(* IEC 61131-3 sources: Jacob-Formschaumtechnik-ISEL-CNC-Retrofit/twincat/PLC/src/4_Machine, 9 files *)

(* ---- FB_Homing.st ---- *)
(* Referenzfahrt als Ablauf: Z zuerst (Spindel nach oben), dann Querachse, dann Portal (Gantry).
   Reihenfolge und Richtung einstellbar (Anforderung 2.2.1). Der Baustein fordert die Fahrt an,
   die Bewegung selbst macht die CNC bzw. der Antrieb. Gantry-Ausrichtung beider Portalseiten
   gehoert in die CNC-Parametrierung. Gruppen: 1 = Z, 2 = X (Quer), 3 = Y (Portal).
   [Annahme] Reihenfolge Z, X, Y, bis Maschinenaufbau bestaetigt.
   Befund 8: Je Gruppe ein Handshake. Erst kommt ein Ruecksetz-Impuls (aResetHomed), dann muss aHomed
   FALSE werden, danach steht bHomeCmd als Pegel, bis aHomed wieder TRUE ist. Zwischen zwei Gruppen
   faellt bHomeCmd mindestens einen Zyklus. Einzelne X/Y-Referenzfahrt nur mit referenziertem Z. *)
FUNCTION_BLOCK FB_Homing
VAR_INPUT
    bStart       : BOOL;                      (* Impuls: alle Achsen in Reihenfolge *)
    aStartAxis   : ARRAY[1..3] OF BOOL;       (* Impuls: nur diese Gruppe *)
    bAbort       : BOOL;
    bHomingOk    : BOOL;
    aHomed       : ARRAY[1..3] OF BOOL;       (* je Gruppe, aus dem einheitlichen Referenzstatus *)
    aOrder       : ARRAY[1..3] OF USINT := [1, 2, 3];
    tTimeout     : TIME := T#120S;
END_VAR
VAR_OUTPUT
    bBusy        : BOOL;
    bDone        : BOOL;
    bError       : BOOL;
    nActiveGroup : USINT;                     (* Gruppe, die gerade referenziert wird, 0 = keine *)
    bHomeCmd     : BOOL;                      (* Anforderung an die CNC/den Antrieb fuer nActiveGroup *)
    aResetHomed  : ARRAY[1..3] OF BOOL;       (* Impuls: Referenzstatus dieser Gruppe loeschen *)
    eHomeState   : ARRAY[1..3] OF E_HomeState;
    nStepOut     : USINT;
END_VAR
VAR
    nStep      : INT;
    nSub       : INT;                         (* 0 Reset senden, 1 auf Reset warten, 2 fahren *)
    nSingle    : USINT;
    rtStart    : R_TRIG;
    rtSingle   : ARRAY[1..3] OF R_TRIG;
    tonTimeout : TON;
    i          : INT;
END_VAR

rtStart(CLK := bStart);
FOR i := 1 TO 3 DO
    rtSingle[i](CLK := aStartAxis[i]);
    aResetHomed[i] := FALSE;
END_FOR
bHomeCmd := FALSE;

IF bAbort OR (bBusy AND NOT bHomingOk) THEN
    IF bBusy AND nActiveGroup > 0 THEN eHomeState[nActiveGroup] := E_HomeState.Open; END_IF
    nStep := 0; nSub := 0; bBusy := FALSE; nActiveGroup := 0; tonTimeout(IN := FALSE);
END_IF

CASE nStep OF
    0:
        IF bHomingOk THEN
            IF rtStart.Q THEN
                bDone := FALSE; bError := FALSE; bBusy := TRUE; nSingle := 0; nStep := 1; nSub := 0;
                FOR i := 1 TO 3 DO eHomeState[i] := E_HomeState.Open; END_FOR
            ELSE
                FOR i := 1 TO 3 DO
                    IF rtSingle[i].Q AND NOT bBusy THEN
                        IF i > 1 AND NOT aHomed[1] THEN
                            bError := TRUE;    (* Z muss zuerst referenziert sein *)
                        ELSE
                            bDone := FALSE; bError := FALSE; bBusy := TRUE; nSingle := TO_USINT(i);
                            nStep := 1; nSub := 0;
                            eHomeState[i] := E_HomeState.Open;
                        END_IF
                    END_IF
                END_FOR
            END_IF
        END_IF
    1, 2, 3:
        IF nSingle > 0 THEN
            nActiveGroup := nSingle;
        ELSE
            nActiveGroup := aOrder[nStep];
        END_IF
        tonTimeout(IN := TRUE, PT := tTimeout);
        CASE nSub OF
            0:  aResetHomed[nActiveGroup] := TRUE;
                eHomeState[nActiveGroup] := E_HomeState.Running;
                nSub := 1;
            1:  IF NOT aHomed[nActiveGroup] THEN nSub := 2; END_IF
            2:  bHomeCmd := TRUE;
                IF aHomed[nActiveGroup] THEN
                    eHomeState[nActiveGroup] := E_HomeState.Done;
                    tonTimeout(IN := FALSE);
                    nSub := 0;
                    IF nSingle > 0 THEN nStep := 4; ELSE nStep := nStep + 1; END_IF
                END_IF
        END_CASE
        IF tonTimeout.Q THEN
            eHomeState[nActiveGroup] := E_HomeState.Error;
            bError := TRUE; bBusy := FALSE; nActiveGroup := 0; nStep := 0; nSub := 0;
            tonTimeout(IN := FALSE);
        END_IF
    4:
        bDone := TRUE; bBusy := FALSE; nActiveGroup := 0; nStep := 0; nSub := 0;
END_CASE
nStepOut := TO_USINT(nStep);
END_FUNCTION_BLOCK

(* ---- FB_Interlocks.st ---- *)
(* Verriegelungsmatrix. Reine Logik ohne Hardwarebezug, daher voll testbar.
   Jede Zeile haengt an einer Anforderung aus der Funktionsliste (Platzhalter-IDs bis Lastenheft da ist). *)
FUNCTION_BLOCK FB_Interlocks
VAR_INPUT
    eMode          : E_OpMode;
    eState         : E_MachState;
    bSafetyOk      : BOOL;
    bAllHomed      : BOOL;
    bDrivesEnabled : BOOL;
    bHmiLinkOk     : BOOL;
    bAnyR2OrHigher : BOOL;
    bAnyR3OrHigher : BOOL;
    bAirOk         : BOOL;
    bHomingBusy    : BOOL;      (* Referenzfahrt laeuft (Befund 8c) *)
    bLimitFreeRun  : BOOL;      (* nur Endschalter-R3 aktiv, Freifahren erlaubt (Befund 15) *)
END_VAR
VAR_OUTPUT
    bProgramStartOk : BOOL;   (* Auto: Start erlaubt *)
    bJogOk          : BOOL;   (* Tippen erlaubt *)
    bHomingOk       : BOOL;
    bSpindleOk      : BOOL;   (* Spindel darf laufen *)
    bAuxOk          : BOOL;   (* Absaugung, Blasluft, Vakuum von Hand *)
    bModeChangeOk   : BOOL;   (* Wechsel nur ohne aktives Programm *)
END_VAR

bProgramStartOk := eMode = E_OpMode.Auto OR eMode = E_OpMode.Setup;
bProgramStartOk := bProgramStartOk AND bSafetyOk AND bDrivesEnabled AND bAllHomed
                   AND NOT bAnyR2OrHigher AND bAirOk AND eState <> E_MachState.Execute AND NOT bHomingBusy;

bJogOk := eMode = E_OpMode.Hand AND bSafetyOk AND bDrivesEnabled AND bHmiLinkOk
          AND (NOT bAnyR3OrHigher OR bLimitFreeRun) AND eState <> E_MachState.Execute AND NOT bHomingBusy;

(* Referenzfahrt nur in Hand und nur im Zustand Idle (nicht in Held/Execute) *)
bHomingOk := eMode = E_OpMode.Hand AND bSafetyOk AND bDrivesEnabled AND NOT bAnyR3OrHigher AND eState = E_MachState.Idle;

bSpindleOk := bSafetyOk AND NOT bAnyR3OrHigher AND eMode <> E_OpMode.Setup;

bAuxOk := bSafetyOk AND eState <> E_MachState.EStop;

bModeChangeOk := eState <> E_MachState.Execute AND eState <> E_MachState.Held;
END_FUNCTION_BLOCK

(* ---- FB_Jog.st ---- *)
(* Tippbetrieb aus der HMI (Anforderungen 2.3.1 und 2.3.2). Nur mit Lebenszeichen der HMI, nur
   in Betriebsart Hand. Befund 6 der Papierpruefung: Tippen startet nur mit einer steigenden Flanke
   der Taste, waehrend alle Freigaben bestehen. Eine beim Wiederkehren der Freigabe (Quittierung,
   Sicherheitskreis, HMI-Lebenszeichen) noch gehaltene Taste startet nichts. Die Achsnummer wird
   beim Start festgehalten. Die Bewegung selbst fordert die CNC an. *)
FUNCTION_BLOCK FB_Jog
VAR_INPUT
    bJogOk       : BOOL;      (* aus FB_Interlocks *)
    bPlus        : BOOL;
    bMinus       : BOOL;
    nAxis        : USINT;     (* 1=X, 2=Y, 3=Z *)
    bRapid       : BOOL;
    nHeartbeat   : UINT;
    tHmiTimeout  : TIME;
    bPlusBlocked  : BOOL;     (* G-01: Endschalter Plus-Seite der gewaehlten Achse ausgeloest, Tippen+ gesperrt *)
    bMinusBlocked : BOOL;     (* Minus-Seite ausgeloest, Tippen- gesperrt *)
END_VAR
VAR_OUTPUT
    bJogPlusReq  : BOOL;
    bJogMinusReq : BOOL;
    nAxisReq     : USINT;
    bRapidReq    : BOOL;
    bHmiLinkOk   : BOOL;
END_VAR
VAR
    nLastHb   : UINT;
    tonLink   : TON;
    rtPlus    : R_TRIG;
    rtMinus   : R_TRIG;
    bActPlus  : BOOL;
    bActMinus : BOOL;
    nAxisLatch: USINT;
    bOkNow    : BOOL;
    nAxisPrev : USINT;
    nStableCyc: USINT;        (* Zyklen, seit denen nAxis unveraendert ist (Befund 16) *)
    bPendPlus : BOOL;         (* Flanke gesehen, wartet auf stabile Achsnummer *)
    bPendMinus: BOOL;
END_VAR

(* Lebenszeichen: Aenderung innerhalb tHmiTimeout *)
IF nHeartbeat <> nLastHb THEN
    nLastHb := nHeartbeat;
    tonLink(IN := FALSE);
END_IF
tonLink(IN := TRUE, PT := tHmiTimeout);
bHmiLinkOk := NOT tonLink.Q AND tHmiTimeout > T#0S;

rtPlus(CLK := bPlus);
rtMinus(CLK := bMinus);
bOkNow := bJogOk AND bHmiLinkOk AND nAxis >= 1 AND nAxis <= 3;

(* Befund 16: Achsnummer und Taste kommen als getrennte ADS-Schreibzugriffe. Start erst, wenn nAxis
   mindestens 2 Zyklen stabil ist; Achswechsel waehrend der Fahrt stoppt sofort. *)
IF nAxis <> nAxisPrev THEN
    nAxisPrev := nAxis; nStableCyc := 0;
ELSIF nStableCyc < 255 THEN
    nStableCyc := nStableCyc + 1;
END_IF

IF NOT bOkNow THEN
    bActPlus := FALSE; bActMinus := FALSE; bPendPlus := FALSE; bPendMinus := FALSE;
ELSE
    (* G-01: Ausgeloester Endschalter beendet das Tippen in dieser Richtung sofort, neue Flanke noetig *)
    IF bPlusBlocked  THEN bActPlus  := FALSE; bPendPlus  := FALSE; END_IF
    IF bMinusBlocked THEN bActMinus := FALSE; bPendMinus := FALSE; END_IF
    IF NOT bPlus  OR bMinus THEN bActPlus  := FALSE; bPendPlus  := FALSE; END_IF
    IF NOT bMinus OR bPlus  THEN bActMinus := FALSE; bPendMinus := FALSE; END_IF
    IF (bActPlus OR bActMinus) AND nAxis <> nAxisLatch THEN
        bActPlus := FALSE; bActMinus := FALSE;
    END_IF
    IF rtPlus.Q  AND NOT bMinus THEN bPendPlus  := TRUE; END_IF
    IF rtMinus.Q AND NOT bPlus  THEN bPendMinus := TRUE; END_IF
    IF bPendPlus AND nStableCyc >= 2 AND NOT bActMinus AND NOT bPlusBlocked THEN
        bActPlus := TRUE; bPendPlus := FALSE; nAxisLatch := nAxis;
    END_IF
    IF bPendMinus AND nStableCyc >= 2 AND NOT bActPlus AND NOT bMinusBlocked THEN
        bActMinus := TRUE; bPendMinus := FALSE; nAxisLatch := nAxis;
    END_IF
END_IF

bJogPlusReq  := bActPlus;
bJogMinusReq := bActMinus;
nAxisReq     := nAxisLatch;
bRapidReq    := bRapid AND (bActPlus OR bActMinus);
END_FUNCTION_BLOCK

(* ---- FB_MachineState.st ---- *)
(* Maschinenzustand. Entscheidet aus Sicherheits- und Meldungsklasse, ob Antriebe freigegeben sind
   und wie reagiert wird. Bewegung und Programm laufen in der CNC, hier nur die Anforderungen.
   Befund 4: Bei NOT-HALT/Tuer/Abbruch/R3/R4 aus Execute oder Held bleibt die Abbruch-Anforderung an die CNC
   als Pegel stehen (bAbortPending), bis die CNC meldet, dass kein Programm mehr aktiv ist. Der NOT-HALT-Zustand
   wird erst danach und nach Quittierung verlassen. *)
FUNCTION_BLOCK FB_MachineState
VAR_INPUT
    bSafetyOk       : BOOL;
    bDrivesAllowed  : BOOL;     (* aus FB_SafetyMonitor *)
    bAnyR2OrHigher  : BOOL;
    bAnyR3OrHigher  : BOOL;
    bAnyR4          : BOOL;
    bAckPending     : BOOL;
    bStartOk        : BOOL;     (* aus FB_Interlocks *)
    bStartCmd       : BOOL;     (* Impuls von der HMI *)
    bHoldCmd        : BOOL;
    bAbortCmd       : BOOL;
    bProgramDone    : BOOL;     (* von der CNC, Flanke genuegt *)
    bProgramActive  : BOOL;     (* von der CNC: Programm laeuft oder Achsen fahren noch *)
    bAck            : BOOL;
    tR4OffDelay     : TIME := T#500MS;   (* Befund 15: Reglerfreigabe faellt bei R4 erst, wenn die CNC steht oder nach dieser Zeit *)
    bDoorOpenAllowed : BOOL;    (* Werkzeugwechsel mit Tuerfreigabe: offene Tuer haelt das Programm an, bricht es nicht ab *)
END_VAR
VAR_OUTPUT
    eState          : E_MachState;
    bEnableDrives   : BOOL;     (* Reglerfreigabe der SPS *)
    bCncStart       : BOOL;     (* Anforderung an die CNC *)
    bCncHold        : BOOL;
    bCncAbort       : BOOL;     (* Pegel, bis die CNC steht *)
    bSpindleStop    : BOOL;     (* Spindel aus, Pegel bei Abbruch/Fehler/NOT-HALT *)
END_VAR
VAR
    rtStart      : R_TRIG;
    rtHold       : R_TRIG;
    rtAbort      : R_TRIG;
    rtAck        : R_TRIG;
    rtDone       : R_TRIG;
    bAbortPending: BOOL;
    ePrev        : E_MachState;
    tonR4Off     : TON;
END_VAR

rtStart(CLK := bStartCmd);
rtHold(CLK := bHoldCmd);
rtAbort(CLK := bAbortCmd);
rtAck(CLK := bAck);
rtDone(CLK := bProgramDone);
bCncStart := FALSE; bCncHold := FALSE; bSpindleStop := FALSE;
ePrev := eState;

(* Vorrang 1: Sicherheitskreis offen -> NOT-HALT-Zustand, Antriebe aus, Programm abbrechen *)
IF NOT bSafetyOk AND bDoorOpenAllowed AND (eState = E_MachState.Execute OR eState = E_MachState.Held) THEN
    (* Werkzeugwechsel bei Spindelstillstand: Tuer offen = Halt, kein Abbruch. Antriebe nimmt die Verdrahtung weg. *)
    IF eState = E_MachState.Execute THEN eState := E_MachState.Held; END_IF
ELSIF NOT bSafetyOk THEN
    IF eState = E_MachState.Execute OR eState = E_MachState.Held THEN
        bAbortPending := TRUE;
    END_IF
    eState := E_MachState.EStop;
ELSIF eState = E_MachState.EStop THEN
    (* Sicherheitskreis wieder zu: Quittierung, Programm muss beendet sein *)
    IF bDrivesAllowed AND rtAck.Q AND NOT bAbortPending THEN eState := E_MachState.Stopped; END_IF
END_IF

(* Vorrang 2: Meldungsklassen *)
IF eState <> E_MachState.EStop THEN
    IF bAnyR4 THEN
        IF eState = E_MachState.Execute OR eState = E_MachState.Held THEN bAbortPending := TRUE; END_IF
        eState := E_MachState.Fault;
    ELSIF bAnyR3OrHigher THEN
        IF eState = E_MachState.Execute OR eState = E_MachState.Held THEN
            bAbortPending := TRUE;
        END_IF
        eState := E_MachState.Aborted;
    ELSIF bAnyR2OrHigher AND eState = E_MachState.Execute THEN
        bCncHold := TRUE;
        eState := E_MachState.Held;
    END_IF
END_IF

(* Normaler Ablauf *)
CASE eState OF
    E_MachState.Stopped:
        IF bDrivesAllowed AND NOT bAnyR3OrHigher AND NOT bAckPending THEN
            eState := E_MachState.Idle;
        END_IF
    E_MachState.Idle:
        IF rtStart.Q AND bStartOk THEN
            bCncStart := TRUE;
            eState := E_MachState.Execute;
        END_IF
    E_MachState.Execute:
        IF rtHold.Q THEN bCncHold := TRUE; eState := E_MachState.Held; END_IF
        IF rtAbort.Q THEN bAbortPending := TRUE; eState := E_MachState.Aborted; END_IF
        IF rtDone.Q THEN eState := E_MachState.Idle; END_IF
    E_MachState.Held:
        IF rtStart.Q AND bStartOk AND NOT bAnyR2OrHigher THEN
            bCncStart := TRUE; eState := E_MachState.Execute;
        END_IF
        IF rtAbort.Q THEN bAbortPending := TRUE; eState := E_MachState.Aborted; END_IF
        IF rtDone.Q THEN eState := E_MachState.Idle; END_IF   (* G-02: Programmende waehrend Halt *)
    E_MachState.Aborted, E_MachState.Fault:
        IF rtAck.Q AND NOT bAnyR3OrHigher AND NOT bAckPending AND NOT bAbortPending THEN eState := E_MachState.Stopped; END_IF
END_CASE

(* G-02: Vorschubhalt als Pegel, solange der Zustand Held ist (ein Ein-Zyklus-Impuls reicht fuer die CNC nicht).
   Er faellt mit dem Fortsetzen (Start) oder Abbruch. [offen] HLI-Semantik bei der Anbindung dokumentieren. *)
IF eState = E_MachState.Held THEN bCncHold := TRUE; END_IF

(* Abbruch bleibt angefordert, bis die CNC steht *)
IF bAbortPending AND NOT bProgramActive AND ePrev = eState AND NOT (rtAbort.Q) THEN
    bAbortPending := FALSE;
END_IF
bCncAbort := bAbortPending;

(* Spindel aus in allen Zustaenden ausser Idle/Execute/Held/Stopped *)
bSpindleStop := bAbortPending OR eState = E_MachState.EStop OR eState = E_MachState.Aborted OR eState = E_MachState.Fault;

(* Befund 15: Bei R4 (Zustand Fault) bremst die CNC gefuehrt (Abbruch laeuft), die Freigabe faellt, sobald
   die CNC kein Programm/keine Bewegung mehr meldet, spaetestens nach tR4OffDelay. NOT-HALT wirkt sofort
   (Sicherheitsrelais nimmt die Freigabe in Hardware, bDrivesAllowed faellt im selben Zyklus). *)
tonR4Off(IN := bAnyR4 OR eState = E_MachState.Fault, PT := tR4OffDelay);
bEnableDrives := bDrivesAllowed AND eState <> E_MachState.EStop
                 AND NOT ((bAnyR4 OR eState = E_MachState.Fault) AND (tonR4Off.Q OR NOT bProgramActive));
END_FUNCTION_BLOCK

(* ---- FB_OpModeManager.st ---- *)
(* Betriebsartenwahl. Wechsel nur im Stillstand (kein Programm, keine Achsbewegung, Spindel steht).
   Ein vorhandener Schluesselschalter (bKeyAuto) hat Vorrang vor der HMI. *)
FUNCTION_BLOCK FB_OpModeManager
VAR_INPUT
    eRequest       : E_OpMode;     (* von der HMI *)
    bStandstill    : BOOL;         (* alle Achsen stehen, Programm nicht aktiv, Spindel steht *)
    bHasKeySwitch  : BOOL;         (* [offen] Schluesselschalter am Pult vorhanden? *)
    bKeyAuto       : BOOL;         (* Schluesselschalter in AUTO *)
END_VAR
VAR_OUTPUT
    eMode          : E_OpMode;
    bChangeBlocked : BOOL;         (* Wunsch abgelehnt, HMI zeigt Hinweis *)
END_VAR

bChangeBlocked := FALSE;

IF bHasKeySwitch AND NOT bKeyAuto AND eRequest = E_OpMode.Auto THEN
    (* Schluessel nicht auf AUTO: Automatik nicht zulaessig *)
    bChangeBlocked := TRUE;
ELSIF eRequest <> eMode THEN
    IF bStandstill THEN
        eMode := eRequest;
    ELSE
        bChangeBlocked := TRUE;
    END_IF
END_IF

(* Schluessel weg von AUTO: sofort zurueck in Hand, sobald Stillstand *)
IF bHasKeySwitch AND NOT bKeyAuto AND eMode = E_OpMode.Auto AND bStandstill THEN
    eMode := E_OpMode.Hand;
END_IF
END_FUNCTION_BLOCK

(* ---- FB_ParamCheck.st ---- *)
(* Prueft beim Start Maschinen-ID und Softwareversion. Passt etwas nicht, bleibt die Maschine gesperrt
   (Meldung 900, R4). Anforderungen 2.11.4 und 2.11.5. *)
FUNCTION_BLOCK FB_ParamCheck
VAR_INPUT
    nIdExpected   : UINT;
    nIdLoaded     : UINT;
    sVerExpected  : STRING(15);
    sVerRunning   : STRING(15);
    bParamsLoaded : BOOL;
END_VAR
VAR_OUTPUT
    bMismatch : BOOL;
END_VAR

bMismatch := NOT bParamsLoaded OR (nIdLoaded <> nIdExpected) OR (sVerExpected <> sVerRunning);
END_FUNCTION_BLOCK

(* ---- FB_ParamInit.st ---- *)
(* Initialisiert die Maschinenparameter und prueft sie auf Plausibilitaet (Befunde 2 und 20).
   Der Parametersatz wird nach der Maschinenkennung des Geraets (GVL_Persistent.nMachineId) gewaehlt,
   damit ein Softwarestand fuer alle Maschinen gilt. Unbekannte Kennung: kein Satz, Maschine gesperrt.
   Uebergangsloesung: Werte stehen hier als Konstanten und entsprechen config/M1.json. Alle Werte ausser
   rSpindleMaxRpm sind Annahmen. Spaeter ersetzt ein Lader (Tc3_JsonXml) die Zuweisungen, die Pruefung bleibt.
   bLoaded wird nur TRUE, wenn alle Werte plausibel sind. *)
FUNCTION_BLOCK FB_ParamInit
VAR_INPUT
    nMachineId : UINT;            (* Kennung des Geraets *)
END_VAR
VAR_IN_OUT
    stParams : ST_MachineParams;
END_VAR
VAR_OUTPUT
    bLoaded  : BOOL;
    bInvalid : BOOL;
    bUnknownId : BOOL;            (* keine Parameter fuer diese Kennung *)
END_VAR
VAR
    bDone     : BOOL;
    nIdLoaded : UINT;
END_VAR

(* Neu laden, wenn sich die Kennung aendert (Inbetriebnahme) *)
IF bDone AND nMachineId <> nIdLoaded THEN bDone := FALSE; END_IF

IF NOT bDone THEN
    bDone := TRUE;
    nIdLoaded := nMachineId;
    bUnknownId := FALSE;
    CASE nMachineId OF
        1:  (* M1 *)
            stParams.nMachineId         := 1;
            stParams.sSwVersionExpected := '0.12.0';   (* Platzhalter, gleiche Quelle wie GVL_Config.sSwVersion: Pruefung wirkt erst mit externem Parametersatz *)
            stParams.eDriveVariant      := E_DriveVariant.Simulation;   (* [offen] bis Antriebsabbildung steht *)
            stParams.nNumAxes           := 4;
            stParams.nNumCncAxes        := 3;
            stParams.rSpindleMaxRpm     := 16600.0;
            stParams.rSpindleMinRpm     := 0.0;
            stParams.rSpindleVoltMax    := 10.0;
            stParams.tSpindleRunUp      := T#8S;
            stParams.tSpindleStandstill := T#10S;
            stParams.tHmiTimeout        := T#500MS;
            stParams.tFeedbackTimeout   := T#3S;
            stParams.bAirMonitoring     := TRUE;
            stParams.bHasToolChanger    := FALSE;
    ELSE
        bUnknownId := TRUE;
        stParams.nMachineId := 0;
    END_CASE
END_IF

bInvalid := bUnknownId OR stParams.rSpindleMaxRpm <= 0.0 OR stParams.rSpindleVoltMax <= 0.0
            OR stParams.tSpindleRunUp <= T#0S OR stParams.tSpindleStandstill <= T#0S
            OR stParams.tHmiTimeout <= T#0S OR stParams.tFeedbackTimeout <= T#0S
            OR stParams.rSpindleMinRpm < 0.0 OR stParams.rSpindleMinRpm >= stParams.rSpindleMaxRpm
            OR stParams.nNumAxes <> 4 OR stParams.nNumCncAxes <> 3
            OR stParams.eDriveVariant <> GVL_Config.eDriveVariant;
bLoaded := bDone AND NOT bInvalid;
END_FUNCTION_BLOCK

(* ---- FB_SafetyMonitor.st ---- *)
(* Liest den Status der festen Sicherheitsverdrahtung (Pilz-Relais, Tuerkontakt) und bildet
   die SPS-Seite der Antriebsfreigabe. Die SPS kann nur zusaetzlich sperren, nie freigeben,
   was das Relais sperrt. Das ist KEINE Sicherheitsfunktion im Sinne ISO 13849.
   Ruhestromprinzip: FALSE = Sicherheitskreis offen. *)
FUNCTION_BLOCK FB_SafetyMonitor
VAR_INPUT
    bRelayFeedbackOk : BOOL;   (* Rueckmeldekontakt Sicherheitsrelais *)
    bDoorClosed      : BOOL;   (* Statussignal Tuer *)
    bFieldbusOk      : BOOL;
    bAck             : BOOL;   (* Quittierung, Impuls *)
    bAirOk           : BOOL;
END_VAR
VAR_OUTPUT
    bSafetyOk     : BOOL;      (* Sicherheitskreis geschlossen *)
    bDrivesAllowed: BOOL;      (* SPS-Freigabe der Antriebe, nur mit Quittierung nach Ausloesung *)
    bLatched      : BOOL := TRUE;   (* Wiederanlauf wartet auf Quittierung; nach dem Anlauf immer TRUE (Befund 7) *)
END_VAR
VAR
    rtAck       : R_TRIG;
    bWasOk      : BOOL;
END_VAR

rtAck(CLK := bAck);
(* Befund 19: Feldbusausfall zaehlt als offener Sicherheitskreis (Eingaenge koennten auf dem letzten Wert stehen) *)
bSafetyOk := bRelayFeedbackOk AND bDoorClosed AND bFieldbusOk;

IF NOT bSafetyOk OR NOT bFieldbusOk THEN
    bLatched := TRUE;           (* Wiederanlauf nie automatisch *)
END_IF
IF bLatched AND bSafetyOk AND bFieldbusOk AND rtAck.Q THEN
    bLatched := FALSE;
END_IF

bDrivesAllowed := bSafetyOk AND bFieldbusOk AND NOT bLatched;
END_FUNCTION_BLOCK

(* ---- FB_ToolChange.st ---- *)
(* Manueller Werkzeugwechsel (Anforderung 2.6.2). M6 mit Werkzeugnummer: Spindel aus, Aufforderung
   am Panel, Programm wartet auf Quittung. Kein Werkzeugwechsler im Umfang (offen: "SW"). *)
FUNCTION_BLOCK FB_ToolChange
VAR_INPUT
    bM6Request   : BOOL;      (* aus FB_MFunctions *)
    nToolNo      : UINT;      (* angeforderte Werkzeugnummer aus der CNC *)
    bSpindleStopped : BOOL;
    bConfirm     : BOOL;      (* Impuls HMI: Wechsel erledigt *)
    bAbort       : BOOL;
END_VAR
VAR_OUTPUT
    bRequest     : BOOL;      (* Aufforderung am Panel *)
    nRequestedTool : UINT;
    bHoldProgram : BOOL;      (* CNC wartet, bis quittiert *)
    bSpindleLock : BOOL;      (* Spindel gesperrt waehrend Wechsel *)
    bDoorRelease : BOOL;      (* Tuer darf geoeffnet werden: Werkzeugwechsel angefordert und Spindel steht. Eine offene Tuer bricht dann das Programm nicht ab. *)
END_VAR
VAR
    rtM6 : R_TRIG;
    rtConfirm : R_TRIG;
END_VAR

rtM6(CLK := bM6Request);
rtConfirm(CLK := bConfirm);

IF rtM6.Q THEN
    bRequest := TRUE; nRequestedTool := nToolNo;
END_IF
bHoldProgram := bRequest;
bSpindleLock := bRequest;
IF bRequest AND ((rtConfirm.Q AND bSpindleStopped) OR bAbort) THEN
    bRequest := FALSE;
END_IF

(* Tuerfreigabe fuer den Werkzeugwechsel: erst bei Spindelstillstand. Die Abschaltung der Antriebe macht weiter die
   feste Verdrahtung (Pilz). Die SPS entscheidet nur zwischen Halt (Wechsel) und Abbruch. [offen] Risikobeurteilung:
   Zustimmtaster, Schluesselschalter, sichere Spindelstillstandsueberwachung. *)
bDoorRelease := bRequest AND bSpindleStopped;
END_FUNCTION_BLOCK
